(* IEC 61131-3 sources: llm-plc-st-eval/data/definitivo/claude-sonnet-4-6/C3/few_shot, 3 files *)

(* ---- ejec_1.st ---- *)
```pascal
PROGRAM PRG_Conversion
VAR_INPUT
    btnMarcha : BOOL; (* Contacto NA: arranque *)
    btnParo   : BOOL; (* Contacto NC: paro *)
END_VAR
VAR_OUTPUT
    motor   : BOOL; (* Bobina motor / contacto de enclavamiento *)
    lampara : BOOL; (* Bobina lámpara *)
END_VAR
VAR
    T1 : TON; (* Temporizador retardo a la conexión *)
END_VAR

(* Rama 1: (btnMarcha OR motor) AND NOT btnParo -> bobina motor *)
(* El contacto NA motor actúa como enclavamiento (auto-retención)  *)
motor := (btnMarcha OR motor) AND NOT btnParo;

(* Rama 2: contacto NA motor habilita el temporizador T1 (PT = 10 s) *)
T1(IN := motor, PT := T#10S);

(* Rama 3: contacto NA T1.Q -> bobina lámpara *)
lampara := T1.Q;

END_PROGRAM
```

(* ---- ejec_2.st ---- *)
```pascal
PROGRAM PRG_Conversion
VAR_INPUT
    btnMarcha : BOOL; (* Contacto NA: arranque *)
    btnParo   : BOOL; (* Contacto NC: paro *)
END_VAR
VAR_OUTPUT
    motor   : BOOL; (* Bobina motor / contacto de enclavamiento *)
    lampara : BOOL; (* Bobina lampara *)
END_VAR
VAR
    T1 : TON; (* Temporizador on-delay, PT = 10 s *)
END_VAR

(* Rama 1: (btnMarcha OR motor) AND NOT btnParo -> bobina motor *)
(* El contacto NA motor actua como enclavamiento (seal-in) *)
motor := (btnMarcha OR motor) AND NOT btnParo;

(* Rama 2: contacto NA motor habilita el temporizador T1 *)
(* Cuando motor se desactiva, T1 se resetea automaticamente *)
T1(IN := motor, PT := T#10S);

(* Rama 3: contacto NA T1.Q -> bobina lampara *)
(* La lampara se enciende cuando el motor lleva 10 s activo *)
lampara := T1.Q;

END_PROGRAM
```

(* ---- ejec_3.st ---- *)
```pascal
PROGRAM PRG_Conversion
VAR_INPUT
    btnMarcha : BOOL; (* Contacto NA: arranque *)
    btnParo   : BOOL; (* Contacto NC: paro *)
END_VAR
VAR_OUTPUT
    motor   : BOOL; (* Bobina motor / contacto de enclavamiento *)
    lampara : BOOL; (* Bobina lampara *)
END_VAR
VAR
    T1 : TON; (* Temporizador, tiempo preestablecido 10 s *)
END_VAR

(* Rama 1: (btnMarcha OR motor) AND NOT btnParo -> bobina motor *)
(* Paralelo = OR, serie = AND, contacto NC = NOT *)
motor := (btnMarcha OR motor) AND NOT btnParo;

(* Rama 2: contacto NA motor habilita el temporizador TON T1 *)
T1(IN := motor, PT := T#10S);

(* Rama 3: contacto NA T1.Q alimenta la bobina lampara *)
lampara := T1.Q;

END_PROGRAM
```
